{attribute 'qualified_only'}
{attribute 'strict'}
TYPE E_ErrorPiton :
(
	No_piston_error							:=0,
	Wating_for_sensor_open_at_Open_cmd		:=1,
	Wating_for_sensor_close_at_Open_cmd		:=2,
	Wating_for_sensor_close_at_Close_cmd	:=3,
	Wating_for_sensor_open_at_Close_cmd		:=4,
	No_status								:=5,
	No_valve_Operation						:=6,
	Error_not_difined						:=9);
END_TYPE

(* stored: Version 1.1.0.1, ProductVersion 3.1.4024.12
   DUT E_ErrorPiton: Id {8e9a8b2f-e58e-4d43-91a5-3920cdc415e1} *)
